Staubli VAL3: init.pgx

public program init()
begin
  // if rs:bReloadIO
  call linkIO(rs:sBusUsing)
  rs:bReloadIO=false
  rs:libSave()
  //  endIf
  //call linkStatusIO()
end
